(* IEC 61131-3 sources: avi-aoi-management/scripts/ai-eval/ngau-nhien/kho/st-tv3-nhap-nhay/mau/src, 1 file *)

(* ---- NhapNhay.st ---- *)
FUNCTION_BLOCK NhapNhay
VAR_INPUT
    BAT : BOOL;
    T_SANG : TIME;
    T_TOI : TIME;
END_VAR
VAR_OUTPUT
    DEN : BOOL;
END_VAR
VAR
    tg : TON;
    toi : BOOL;   (* đang ở pha tối *)
END_VAR
    IF NOT BAT THEN
        toi := FALSE;
        tg(IN := FALSE);
    ELSE
        IF toi THEN
            tg(IN := TRUE, PT := T_TOI);
        ELSE
            tg(IN := TRUE, PT := T_SANG);
        END_IF
        IF tg.Q THEN
            (* đổi pha; mốc pha mới = chu kỳ này *)
            toi := NOT toi;
            tg(IN := FALSE);
            IF toi THEN
                tg(IN := TRUE, PT := T_TOI);
            ELSE
                tg(IN := TRUE, PT := T_SANG);
            END_IF
        END_IF
    END_IF
    DEN := BAT AND NOT toi;
END_FUNCTION_BLOCK
